PROGRAM TC3_Examples
VAR
	bOnlyRunOnce : BOOL;
	
	// Variables used to show how functions can operate
	fFarenheit : REAL;
	
	nReturnGreater : INT;
	nReturnSmaller : INT;
	
	nNumA : INT;
	nNumB : INT;
	
END_VAR

IF NOT bOnlyRunOnce THEN
	Tc2_System.ADSLOGSTR(msgCtrlMask := Tc2_System.Global_Variables.ADSLOG_MSGTYPE_ERROR OR Tc2_System.Global_Variables.ADSLOG_MSGTYPE_LOG,
						msgFmtStr := 'Hello World!',
						strArg := '');
	bOnlyRunOnce := TRUE;
END_IF

fFarenheit := Celsius_To_Farenheit(fCelsius := 5.0);

Greater_Smaller(nNumber1 := 2, nNumber2 := 9, nGreater => nReturnGreater, nSmaller => nReturnSmaller);

SwapNums(nNumA, nNumB);

POU();

END_PROGRAM

(* stored: Version 1.1.0.1
   POU TC3_Examples: Id {79d2776d-afee-479b-9286-cbec8c87fd10}, SpecialFunc None *)
